FUNCTION_BLOCK RoboStation (* Composite Function Block Type *)
  (* Standard: 61499-2 *)
  (* Version 0.0, 7/2/2026, template *)
  PACKAGE Main;
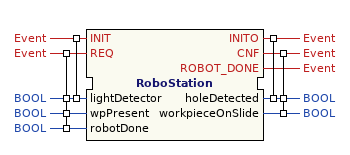
  EVENT_INPUT
    INIT WITH lightDetector; (* Initialization Request *)
    REQ WITH lightDetector, wpPresent, robotDone; (* Normal Execution Request *)
  END_EVENT
  EVENT_OUTPUT
    INITO WITH holeDetected; (* Initialization Confirm *)
    CNF WITH holeDetected, workpieceOnSlide; (* Execution Confirmation *)
    ROBOT_DONE;
  END_EVENT
  VAR_INPUT
    lightDetector : BOOL; (* Input event qualifier *)
    wpPresent : BOOL;
    robotDone : BOOL;
  END_VAR
  VAR_OUTPUT
    holeDetected : BOOL; (* Output event qualifier *)
    workpieceOnSlide : BOOL;
  END_VAR
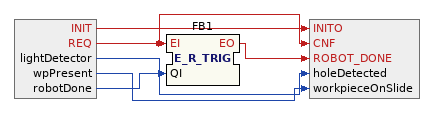
  FBS
    FB1 : E_R_TRIG;
  END_FBS
  EVENT_CONNECTIONS
    REQ TO FB1.EI;
    REQ TO CNF;
    INIT TO INITO;
    FB1.EO TO ROBOT_DONE;
  END_CONNECTIONS
  DATA_CONNECTIONS
    robotDone TO FB1.QI;
    lightDetector TO holeDetected;
    wpPresent TO workpieceOnSlide;
  END_CONNECTIONS
END_FUNCTION_BLOCK
